Fanuc KAREL source: KO00045.KL

PROGRAM KO00045
%NOLOCKGROUP
%ENVIRONMENT MIR
VAR
  P1: POSITION
  P2: JOINTPOS
  F: BOOLEAN
  OUT: POSITION
BEGIN
  F = TRUE
  OUT = MIRROR(P1, P2, F)
END KO00045
